Universal Robots PolyScope program: MainCall.urp

Program MainCall (createdIn=3.0.0 lastSavedIn=3.0.0 directory=/programs installation=default)
Robot Program (runOnlyOnce=true motionType=MoveJ speed=1.047198 acceleration=1.396263 useActiveTCP=false)
  'Program generated by RoboDK v6.0.7 for ABB IRB 120-3/0.6 on XX/XX/XXXX 18:00:00'
  'Using nominal kinematics.'
  'Using Ref. Frame S: p[1.234570, -0.098765, 0.050500, 0.000000, 0.000000, 0.523599]'
  Script: movej([0.000000, -0.174533, 0.349066, 0.000000, 0.523599, 0.000000],1.20000,0.75000,0,0.0000)
  MoveJ speed 42.97 deg/s, acceleration 68.75 deg/s^2 (useActiveTCP=true)
    Waypoint Waypoint_1: TCP in base x=426.318 y=20 z=422.034 mm, rx=0.1383 ry=2.2532 rz=-0.2966 rad; joints [0, -10, 20, 0, 30, 0] deg
  Call SubProg2
  Call NotAProgram
SubProgram  [hidden by the author, left out]
SubProgram  [hidden by the author, left out]
SubProgram SubProg2 [hidden by the author, left out]
SubProgram NotAProgram [hidden by the author, left out]
